Fanuc KAREL source: kt00082.KL

-- PROVISIONAL review KL for V1013-1; original PC SHA256 8c34715a99e22263f4d4c612ef6246c21be561dda751410901ec3df4c98f8179
-- Incomplete behavior may be omitted. Consult companion uncertainty JSON. Do not deploy.
PROGRAM KT00082
%NOLOCKGROUP
VAR
  I2 : INTEGER
  OUT : REAL
-- UNRESOLVED_DECL Y1 type=002018
BEGIN
  -- UNRESOLVED_PC offsets 5-19; opcodes 2E,22,9D,33,B2
  -- UNRESOLVED_PC offsets 24-35; opcodes 2E,23
  -- UNRESOLVED_PC offsets 40-63; opcodes 22,9D,33,B1,21,54,64,23
  -- UNRESOLVED_PC offsets 68-72; opcodes 7F
END KT00082
